Fanuc KAREL source: kt00903.KL

-- PROVISIONAL review KL for V1013-1; original PC SHA256 0a8362d9b30230f2e6650aa8d2a49d0fde803e2953f5bf7ad19dfa1506fb4d32
-- Incomplete behavior may be omitted. Consult companion uncertainty JSON. Do not deploy.
PROGRAM KT00903
%NOLOCKGROUP
BEGIN
  -- UNRESOLVED_PC offsets 5-28; opcodes 27,22,1C,31,4A
  -- UNRESOLVED_PC offsets 33-37; opcodes 7F
END KT00903
